Fanuc KAREL source: kb00049.KL

PROGRAM KB00049
%STACKSIZE=65535
%PRIORITY=65535
%NOLOCKGROUP
VAR
P1 : STRING[80]
P2 : INTEGER
P3 : INTEGER
BEGIN
P1='A'
P2=1
P3=1
CREATE_TPE(P1,P2,P3)
END KB00049
